Fanuc KAREL source: KB00166.KL

PROGRAM KB00166
%NOLOCKGROUP
%ENVIRONMENT REGOPE
VAR
  P1: INTEGER
  P2: JOINTPOS
  P3: INTEGER
BEGIN
  P1 = 1
  P3 = 1
  SET_JPOS_REG(P1, P2, P3)
END KB00166
